Fanuc KAREL source: KC00037.KL

PROGRAM KC00037
%NOLOCKGROUP
%ENVIRONMENT UIF
VAR
  I: INTEGER
  J: INTEGER
  K: INTEGER
  R: REAL
  B: BOOLEAN
  S: STRING[80]
  T: STRING[80]
  P: PATH
  Q: PATH
  AI: ARRAY[8] OF INTEGER
  AB: ARRAY[244] OF BYTE
BEGIN
  CHECK_DICT(S,I,J)
END KC00037
